(* IEC 61131-3 sources: P26002_Bosch_HDPump/P26002_Bosch_HDPump_PLC, 7 files *)

(* ---- CAN_Signals.gvl ---- *)
VAR_GLOBAL

(* ======================================================================== *)
    (* 4. Lokale Prozessvariablen für ALLE gelesenen Messwerte (Rx)             *)
    (* ======================================================================== *)
    rTecu_cpu                   : REAL; (* ID 16#456: ECU CPU Temperatur *)
    rPrail_nom                  : REAL; (* ID 16#650: Fuel pressure HP - set point *)
    rTfuel                      : REAL; (* ID 16#650: Fuel temperature HP *)
    rToil                       : REAL; (* ID 16#650: Öltemperatur *)
    rPrail_650                  : REAL; (* ID 16#650: Fuel pressure HP - side 1 *)
    rMsv_divy_angle             : REAL; (* ID 16#660: MSV Förderwinkel *)
    rAngle_eng_hdp              : REAL; (* ID 16#660: Motorwinkel HDP Messung *)
    rTinj                       : REAL; (* ID 16#660: Einspritzdauer *)
    rPrail_660                  : REAL; (* ID 16#660: Fuel pressure HP - side 2 *)
    rTekp                       : REAL; (* ID 16#670: Fuel temp after low press pump *)
    rPekp                       : REAL; (* ID 16#670: Fuel press after low press pump *)
    rPfuel                      : REAL; (* ID 16#670: Kraftstoffdruck *)
    rEngine_RPM                 : REAL; (* ID 16#680: Drehzahl / RPM *)

    (* ======================================================================== *)
    (* 5. Lokale Variablen für die zu SCHREIBENDEN Werte (Tx)                   *)
    (* ======================================================================== *)
    (* ID 16#700 *)
    rWrite_Set_RPM              : REAL  := 2500.0;
    rWrite_Actual_RPM           : REAL  := 2498.0;
    bWrite_valid_RPM            : BOOL  := TRUE;

    (* ID 16#710 *)
    rWrite_Oil_pressure         : REAL  := 4.5;    (* bar *)
    rWrite_Oil_temperature      : REAL  := 85.0;   (* °C *)
    bWrite_Oil_pressure_OK      : BOOL  := TRUE;
    bWrite_Oil_temperature_OK   : BOOL  := TRUE;

    (* ID 16#720 *)
    rWrite_Fuel_temperature     : REAL  := 25.0;   (* °C *)
    rWrite_Fuel_supply_pressure : REAL  := 5.0;    (* bar *)
    bWrite_Fuel_temperature_OK  : BOOL  := TRUE;
    bWrite_Fuel_supply_press_OK : BOOL  := TRUE;

    (* ID 16#730 *)
    rWrite_Fuel_Mass_Flow_1     : REAL  := 12.5;   (* kg/h *)
    rWrite_Fuel_Mass_Flow_2     : REAL  := 12.4;
    rWrite_Fuel_Mass_Flow_3     : REAL  := 0.0;
    bWrite_valid_Fuel_Mass_Flow : BOOL  := TRUE;

    (* ID 16#800 *)
    wWrite_ERROR_Bits           : WORD  := 16#0000;

    (* ID 16#900 *)
    nWrite_Counter_LAP          : USINT := 1;
    nWrite_Counter_FREE_TRIGGER : USINT := 0;

    (* ID 16#910 (reserviert) *)
    wWrite_RPM_Profile          : WORD  := 16#0000;

END_VAR

(* ---- GlobalVariables.gvl ---- *)
VAR_GLOBAL
system : System;
req_EmgStop_bySoftware : BOOL := FALSE;
reset_EmgStop : BOOL := FALSE;

User : User_InOut;
OP_List: ARRAY[0..10] OF OPoint;

Thermostat : Thermostat;
OilConditioning : OilConditioning;
FuelSupply : FuelSupply;

AutomaticOperation : FB_AutomaticOperation;
fbThermostat: FB_Thermostat;
fbOilConditionin: FB_OilConditioning;
fbFuelSupply: FB_FuelSupply;

HW_DI_ECU_RUNNING : BOOL; (* Kanal entsprechend benennen! *)
END_VAR

VAR_GLOBAL RETAIN
	Retain_Settings : UserSettings;
END_VAR

(* ---- FB_AutomaticOperation.st ---- *)
FUNCTION_BLOCK FB_AutomaticOperation
VAR_INPUT
	system_state : System;
	Enable  : BOOL;
    Stop    : BOOL;
    Reset   : BOOL;
    sequence_active : BOOL;

    coldStart_oil_pressure: REAL := 1.8; (* bar *)
	coldStart_oil_min_tempterature: REAL := 50; (* °C *)
	coldStart_fuelsupply_pressure: REAL := 2; (* bar *)
	coldStart_fuelsupply_min_tempterature: REAL := 50; (* °C *)
	coldStart_RPM_settings: REAL := 2000;

	normalOperation_oil_pressure: REAL := 2.5;(* bar *)
END_VAR

VAR_OUTPUT
	State   : state_op_manager; (* OP_Settle und OP_Hold brauchen wir in diesem Projekt nicht *)
    Busy    : BOOL;
    Done    : BOOL;
    Error   : BOOL;
    ErrMsg	: STRING(255);

    (* ----------------------------- *)
	(* ----- Sequence Control ------ *)
	(* ----------------------------- *)

    start_sequence: BOOL;
    stop_sequence: BOOL;
    coldStart_RPM : REAL;

     (* --- Konfiguration --- *)
    current_OP: OPoint;

END_VAR

VAR_IN_OUT
	IO_User : User_InOut;
	IO_Thermostat : Thermostat;
	IO_OilConditioning: OilConditioning;
	IO_FuelSupply: FuelSupply;
	IO_GlobalOP_List : ARRAY[0..10] OF OPoint;
END_VAR

VAR
	NextState  : state_op_manager;
    LastState  : state_op_manager;

    rpm_rampup: FB_RampTON;
    rpm_rampup_time: TIME := T#2m;
    rpm_rampup_Done: BOOL;

    prep_settle_timer: TON;
    prep_settle_time: TIME := T#60s;

	bEntry			: BOOL := TRUE;
	bInitDone       : BOOL := FALSE;
END_VAR

(* ----------------------------- *)
(* -------- Enable-Gate -------- *)
(* ----------------------------- *)
IF NOT Enable OR system_state.state = SYS_ERROR OR system_state.state = SYS_STANDBY THEN
	bInitDone := FALSE;
    State     := OP_INIT;
    LastState := OP_INIT;
    Busy      := FALSE;
    Done      := FALSE;
    Error     := FALSE;
    IO_User.Input.start := FALSE;
    RETURN;
END_IF;

(* ------------------------------------------------ *)
(* Default assignments                              *)
(* ------------------------------------------------ *)
NextState := State;
Busy  := FALSE;
Done  := FALSE;
Error := FALSE;
coldStart_RPM := 0.0;
rpm_rampup.bExecute := FALSE;
IO_Thermostat.enable := FALSE;
IO_OilConditioning.enable := FALSE;
IO_FuelSupply.enable := FALSE;

(* ------------------------------------------------ *)
(* Entry-Erkennung                                  *)
(* ------------------------------------------------ *)
bEntry := (State <> LastState);

(* ------------------------------------------------ *)
(* State Machine                                    *)
(* ------------------------------------------------ *)
CASE State OF

	OP_INIT:
	    Busy  := FALSE;
		Done  := FALSE;
		Error := FALSE;

	    IF NOT bInitDone THEN

	    ; (* Alle Infos einlesen, ggf Geräte verbinden, Geräte-Status prüfen... *)

	    bInitDone := TRUE;
	    END_IF

	    IF bInitDone THEN
	        NextState := OP_IDLE;
	        IO_User.Output.operation_status_msg := 'INFO: OP Manager initialized.';
	    END_IF

    OP_IDLE:
	    Busy  := FALSE;
		Done  := FALSE;
		Error := FALSE;

    	; (* Warten auf neue Startbedingungen *)
    	(* ------------------------------------------ *)
	    (* Startbedingung prüfen                      *)
	    (* ------------------------------------------ *)
	    Act_CheckStartConditions;

    OP_PREP:
    	Busy := TRUE;
	    Done := FALSE;
	    Error := FALSE;

	    IO_Thermostat.enable := TRUE;
		IO_OilConditioning.enable := TRUE;
		IO_FuelSupply.enable := TRUE;

	    (* Thermostat an *)
	    IO_Thermostat.target_setpoint := current_OP.Fuel_temperature;
	    IO_Thermostat.start := TRUE;

	    (* Ölkonditionierung an *)
	    IF (IO_OilConditioning.actualOil_temperature < coldStart_oil_min_tempterature+5) THEN
	    	IO_OilConditioning.setOil_pressure := coldStart_oil_pressure;
	    ELSE
	    	IF current_OP.Oil_pressure > normalOperation_oil_pressure THEN
	    		IO_OilConditioning.setOil_pressure := current_OP.Oil_pressure;
	    	ELSE
	    		IO_OilConditioning.setOil_pressure := normalOperation_oil_pressure; (* Agleich OP-Vorgabe *)
	    	END_IF
	    END_IF

	    IO_OilConditioning.setOil_temperature := current_OP.Oil_temperature; (* Wie bekomme ich die Temperatur ins ÖL? *)

	    IO_OilConditioning.start := TRUE;

	    (* Ramp up RPM *)
	    IF bEntry THEN
	    	rpm_rampup(bExecute := FALSE); (* Einmal zurücksetzen *)
	    ELSE
			rpm_rampup(
			 	bExecute := TRUE,
			 	fStartVal := 0.0,
			 	fTargetVal := coldStart_RPM_settings,
			 	tRampTime := rpm_rampup_time,
			 	fCurrentVal => coldStart_RPM,
			 	bDone => rpm_rampup_Done
			);
		END_IF

	    IF IO_Thermostat.SVreached AND
	    	IO_OilConditioning.pressure_SVreached AND
	    	IO_OilConditioning.temperature_SVreached THEN

	    	prep_settle_timer.IN := TRUE;
	    END_IF

	    IF prep_settle_timer.Q THEN
	    	IO_FuelSupply.SV := current_OP.Fuel_supply_pressure;
	    	IO_FuelSupply.start := TRUE;
	    END_IF

	    IF IO_Thermostat.SVreached AND
	    	IO_OilConditioning.pressure_SVreached AND
	    	IO_OilConditioning.temperature_SVreached AND
	    	IO_FuelSupply.SVreached AND
	    	rpm_rampup_Done THEN

	    	NextState := OP_EXECUTE;
	    END_IF

    OP_EXECUTE:
	    Busy := TRUE;
	    Done := FALSE;
	    Error := FALSE;

	    IO_Thermostat.enable := TRUE;
		IO_OilConditioning.enable := TRUE;
		IO_FuelSupply.enable := TRUE;

	    (* Benzin-Versorgung an*)
	    (* Nockenwellenantrieb nach Drehzahlvorgabe fahren*)

	OP_FINISHED:
	    Busy := FALSE;
	    Done := TRUE;
	    Error := FALSE;

	    IO_Thermostat.enable := TRUE;
		IO_OilConditioning.enable := TRUE;
(*		IO_FuelSupply.enable := TRUE; *)

	    (* Benzin-Versorgung aus *)
	    IO_FuelSupply.stop := TRUE;

	    (* Nockenwellenantrieb aus*)

	    IF IO_User.Input.continuous THEN
	    	Act_CheckStartConditions;
	    ELSE
	    	(*Cooldown: Thermostat aus, Ölkonditionierung aus*);
	    	IO_Thermostat.stop := TRUE;
	    	IO_OilConditioning.stop := TRUE;

	    END_IF

	OP_ERROR_SHUTDOWN:
	    Error := TRUE;
	    Busy := TRUE;

	OP_ERROR:
	    Error := TRUE;
	    Done := TRUE;

END_CASE;

(* ------------------------------------------------ *)
(* Global transitions                               *)
(* ------------------------------------------------ *)
IF IO_User.Input.cancel THEN
    IF State <> OP_INIT AND State <> OP_ERROR THEN
        NextState := OP_FINISHED;
        IO_User.Input.start := FALSE;
        IO_User.Input.continuous := FALSE;
    ELSIF State = OP_ERROR_SHUTDOWN THEN
    	NextState := OP_ERROR;
    	IO_User.Input.start := FALSE;
        IO_User.Input.continuous := FALSE;
    END_IF
END_IF

IF IO_User.Input.skipOP THEN
    IF State <> OP_INIT AND State <> OP_ERROR THEN
        NextState := OP_FINISHED;
        IO_User.Input.start := TRUE;
        IO_User.Input.continuous := TRUE;
    END_IF
END_IF

(* ------------------------------------------------ *)
(* ---------- Subsystem Error Detection ----------- *)
(* ------------------------------------------------ *)

(* FÜR BOSCHPRÜFSTAND: MFC FEHLER, FU Fehler, Validierungs Probleme?*)

(* IF 	(SUBP_MfcControl.ErrorDetected OR *)
(*	SUBP_HeaterControl.ErrorDetected) OR *)
(*	system.ALARM_VORALARM_H2_CT_STBQ1 AND *)
(*	State <> OP_ERROR_SHUTDOWN AND *)
(*	State <> OP_ERROR *)
(* THEN *)
(*			NextState := OP_ERROR_SHUTDOWN; *)
(*			IF SUBP_MfcControl.ErrorDetected THEN *)
(*				ErrMsg := SUBP_MfcControl.ErrMsg; *)
(*			ELSIF SUBP_HeaterControl.ErrorDetected THEN *)
(*				ErrMsg := SUBP_HeaterControl.ErrMsg; *)
(*			ELSIF system.ALARM_VORALARM_H2_CT_STBQ1 THEN *)
(*				ErrMsg := 'H2 Gas PreAlarm > 5% LowerExplosionLimit - ERROR_SHUTDOWN triggered!'; *)
(*			ELSE *)
(*				ErrMsg := 'Unknown Error detected'; *)
(*			END_IF *)
(*			Act_StateUpdate; *)
(*			RETURN; *)
(* END_IF *)

(* ------------------------------------------------ *)
(* --------- Aktualisierung Statemachine ---------- *)
(* ------------------------------------------------ *)

Act_StateUpdate;

 (* ====== PROGRAMM ENDE ====== *)
END_FUNCTION_BLOCK

ACTIONS
	ACTION Act_StateUpdate
		(* ------------------------------------------------ *)
		(* State update                                     *)
		(* ------------------------------------------------ *)
		LastState := State;
		IF NextState <> State THEN
		    State := NextState;
		END_IF;
	END_ACTION

	ACTION Act_CheckStartConditions

		current_OP := IO_GlobalOP_List[1]; (* Aktuell keine OP-Liste unterstützt *)

		IF current_OP.ProfileConfig.bDataReady AND NOT current_OP.processed THEN
			current_OP.ProfileConfig.bProfileValid := TRUE;
			NextState := OP_PREP;
		END_IF

	END_ACTION

END_ACTIONS

(* ---- MAIN.st ---- *)
PROGRAM MAIN

(*
[ ] OP_Execute
[ ] OP_Finished
[ ] FB_Thermostat
[x] FB_OilConditioning
[x] FB_FuelSupply
[ ] VERIFY RPM
[ ] VERIFY FLOW
*)
VAR
next_state : state_system;
last_state : state_system;

(* GLOBAL ERROR HANDLING *)
was_error: BOOL := FALSE;
ErrorDelayTimer : TON;         (* Delay for Error Detection *)
TriggerTime : TIME := T#1s;
ResetTrigger : TP;
StopTrigger : TP;
ALARM_ARRAY: ARRAY [1..20] OF BOOL;
a : INT; (* warnings iterative varibale *)
WARNING_ARRAY: ARRAY [1..30] OF BOOL;
w : INT; (* warnings iterative varibale *)
i : INT; (*Iteration Variable*)

(* Reset Device Errors *)
resetMfCError : BOOL;
resetEvapError : BOOL;

END_VAR

ACT_EmgStop_bySoftware;
ACT_READ_SafetyStatus;
Act_UserOutput;

ACT_StateMachine;

END_PROGRAM

ACTIONS

ACTION ACT_InitSystem
User.Settings := Retain_Settings;
;
END_ACTION

ACTION ACT_StateMachine

(* Defaults *)
AutomaticOperation.Enable := FALSE;
AutomaticOperation.Reset := FALSE;

system.state := next_state;

	CASE system.state OF
		SYS_STANDBY:
						IF system.alarm OR system.error THEN
							next_state := SYS_ERROR;
							RETURN;
						END_IF

						IF NOT system.is_init THEN
							ACT_InitSystem;
							system.is_init := TRUE;
						END_IF;

						IF User.Input.OperationModeReq THEN
							next_state := SYS_AUTO_READY;
						END_IF

		SYS_ERROR :
						ResetTrigger(IN:= User.Input.reset_Error_byUser, PT:= TriggerTime);

						IF  ResetTrigger.Q THEN
							reset_EmgStop := TRUE;
							User.Input.reset_Error_byUser := FALSE;
							AutomaticOperation.Enable := TRUE;
						END_IF

		SYS_AUTO_BUSY,SYS_AUTO_READY :

						IF system.alarm OR system.error THEN
							next_state := SYS_ERROR;
							RETURN;
						END_IF

						IF HW_DI_ECU_RUNNING THEN (* Kanal entsprechend benennen! *)
							AutomaticOperation.Enable := TRUE;
						ELSE
							AutomaticOperation.Enable := FALSE;
							 WARNING_ARRAY[2] := TRUE; (* Warnung: ECU nicht an! Kein Betrieb möglich *)
						END_IF

						IF User.Input.reset_Error_byUser THEN
							AutomaticOperation.Reset := TRUE;
						END_IF

						IF User.Input.StandbyModeReq THEN
							AutomaticOperation.Stop := TRUE;
						END_IF

		SYS_MANUAL :

						IF system.alarm OR system.error THEN
							next_state := SYS_ERROR;
							RETURN;
						END_IF

						IF User.Input.StandbyModeReq THEN
							next_state := SYS_STANDBY;
							RETURN;
						END_IF
		;
	ELSE
		next_state := SYS_ERROR; (* Other States not allowed!!! *)
		system.status_msg := 'ERROR: State Request NOT allowed!';
	END_CASE

AutomaticOperation(
 IO_User := User,
 IO_Thermostat := Thermostat,
 IO_OilConditioning := OilConditioning,
 IO_FuelSupply := FuelSupply,
 IO_GlobalOP_List := OP_List
);
fbThermostat(fbIO_Thermostat := Thermostat);
fbOilConditionin(fbIO_OilConditioning := OilConditioning);
fbFuelSupply(
 	fbIO_FuelSupply := FuelSupply,
 	SupplyFuelPumpPIDsettings := User.Settings.SupplyFuelPumpPIDsettings,
 	SupplyFuelPump_pressure_tolerance := User.Settings.SupplyFuelPump_pressure_tolerance
);

CASE AutomaticOperation.State OF

	OP_PREP, OP_EXECUTE: next_state := SYS_AUTO_BUSY;

	OP_FINISHED: next_state := SYS_STANDBY;

	OP_ERROR_SHUTDOWN, OP_ERROR: WARNING_ARRAY[1] := TRUE; (* Warnung: Automatic Programm in ERROR Condition *)

END_CASE

(* Global User Input Reset *)
User.Input.reset_Error_byUser := FALSE;
User.Input.StandbyModeReq := FALSE;
User.Input.OperationModeReq := FALSE;

last_state := system.state;
END_ACTION

ACTION Act_UserOutput

		Retain_Settings := User.Settings; (* Backup in Retain Variable *)

		User.Output.SystemState := system;

	END_ACTION

ACTION ACT_EmgStop_bySoftware
	StopTrigger(IN:= User.Input.EmgStop_Req_byUser, PT:= TriggerTime);
	req_EmgStop_bySoftware := StopTrigger.Q;

	IF req_EmgStop_bySoftware THEN
		User.Input.EmgStop_Req_byUser := FALSE;
	END_IF
	;
END_ACTION

ACTION ACT_READ_SafetyStatus (* Wird direkt im Safetyprogramm gemappt *)

		ALARM_ARRAY[1] := system.ALARM_SAI_DiagnosticError;
		ALARM_ARRAY[2] := system.ALARM_GASALARM_H2_ST_STBQ2;
		ALARM_ARRAY[3] := system.ALARM_GASALARM_H2_CT_STBQ1;
		ALARM_ARRAY[4] := system.ALARM_NotAusTaster_1_STFS1;
		ALARM_ARRAY[5] := system.ALARM_NotAusTaster_2_BPSF1;
		ALARM_ARRAY[6] := system.ALARM_EmgStop_bySoftware_activated;
		ALARM_ARRAY[7] := system.ALARM_N2Supply_STBP1;
		ALARM_ARRAY[8] := system.ALARM_HeaterLimit_T_STBT1;
		ALARM_ARRAY[9] := system.ALARM_HeaterLimit_T_STBT2;
		ALARM_ARRAY[10] := system.ALARM_NotAusTaster_1_STFS1_Discrepancy;
		ALARM_ARRAY[11] := system.ALARM_NotAusTaster_2_BPSF1_Discrepancy;
		ALARM_ARRAY[12] := system.ALARM_QA1_Discrepancy;
		ALARM_ARRAY[13] := system.ALARM_QA2_Discrepancy;
		ALARM_ARRAY[14] := system.ALARM_Draeger_Fault;

		FOR i:= 1 TO 20 DO
			IF ALARM_ARRAY[i] THEN
				system.alarm := TRUE;
			END_IF
		END_FOR

	END_ACTION

	ACTION ACT_ResetWarnings

	FOR w := 1 TO 30 DO
		WARNING_ARRAY[w] := FALSE;
	END_FOR

	END_ACTION

	ACTION ACT_CAN_COMMUNICATION
		;
	END_ACTION

END_ACTIONS

(* ---- PRG_MS7_CAN_Handler.st ---- *)
(********************************************************************************
 * PROGRAM: PRG_MS7_CAN_Handler
 *
 * Beschreibung:
 *   Erweitertes Anwendungsbeispiel für das Auslesen und Schreiben des
 *   CAN-Netzwerks (Bosch MS7 Logger / ECU) an einer Bachmann M1 Steuerung.
 *
 *   KANAL-ÜBERSICHT:
 *   ----------------------------------------------------------------------------
 *   EMPFANG (R / Rx):
 *     - Kanal 1 (Rx): ID 16#650 (prail_nom, tfuel, toil, prail_650)
 *     - Kanal 2 (Rx): ID 16#660 (msv_divy_angle, angle_eng_hdp, tinj, prail_660)
 *     - Kanal 3 (Rx): ID 16#670 (tEKP, pEKP, pfuel)
 *     - Kanal 4 (Rx): ID 16#456 (tecu_cpu)
 *     - Kanal 5 (Rx): ID 16#680 (Drehzahl / RPM)
 *
 *   SENDEN (W / Tx):
 *     - Kanal 6  (Tx): ID 16#700 (Set RPM, Actual RPM, valid RPM)
 *     - Kanal 7  (Tx): ID 16#710 (Oil pressure, Oil temperature, Status OK-Bits)
 *     - Kanal 8  (Tx): ID 16#720 (Fuel temp, Fuel supply press, Status OK-Bits)
 *     - Kanal 9  (Tx): ID 16#730 (Fuel Mass Flow 1, 2, 3, valid Bit)
 *     - Kanal 10 (Tx): ID 16#800 (ERROR_Bits)
 *     - Kanal 11 (Tx): ID 16#900 (Counter LAP, Counter FREE TRIGGER)
 *     - Kanal 12 (Tx): ID 16#910 (RPM Profile - reserviert)
 ********************************************************************************)
PROGRAM PRG_MS7_CAN_Handler
VAR
    (* ======================================================================== *)
    (* 1. Konfigurationstabelle / Maske aller CAN-Kanäle (Botschaftsebene)      *)
    (* ======================================================================== *)
    canChannels                 : ARRAY [1..32] OF ST_CAN_Broker_Channel;
    bConfigDone                 : BOOL := FALSE;

    (* Hardware CAN-Broker Instanz (modular bis 32 Kanäle) *)
    fbBroker                    : FB_CAN_Broker_Modular;
    bBrokerReady                : BOOL;
    bBrokerError                : BOOL;
    nBrokerErrorID              : DINT;

    (* ======================================================================== *)
    (* 2. Signal-Instanzen zum LESEN (Rx)                                       *)
    (* ======================================================================== *)
    (* Kanal 4: Botschaft 16#456 (1110 dez) *)
    fb_tecu_cpu                 : FB_CAN_Signal;

    (* Kanal 1: Botschaft 16#650 (1616 dez) *)
    fb_prail_nom                : FB_CAN_Signal; (* Fuel press HP - set point (Bit 0, 16 Bit) *)
    fb_tfuel                    : FB_CAN_Signal; (* Fuel temp HP (Bit 16, 8 Bit) *)
    fb_toil                     : FB_CAN_Signal; (* Oil temp (Bit 24, 8 Bit) *)
    fb_prail_650                : FB_CAN_Signal; (* Fuel press HP - side 1 (Bit 48, 16 Bit) *)

    (* Kanal 2: Botschaft 16#660 (1632 dez) *)
    fb_msv_divy_angle           : FB_CAN_Signal;
    fb_angle_eng_hdp            : FB_CAN_Signal;
    fb_tinj                     : FB_CAN_Signal;
    fb_prail_660                : FB_CAN_Signal; (* Fuel press HP - side 2 (Bit 48, 16 Bit) *)

    (* Kanal 3: Botschaft 16#670 (1648 dez) *)
    fb_tEKP                     : FB_CAN_Signal; (* Fuel temp after low press pump (Bit 0, 16 Bit) *)
    fb_pEKP                     : FB_CAN_Signal; (* Fuel press after low press pump (Bit 16, 16 Bit) *)
    fb_pfuel                    : FB_CAN_Signal; (* Fuel pressure (Bit 32, 8 Bit) *)

    (* Kanal 5: Botschaft 16#680 (1664 dez) *)
    fb_engine_RPM               : FB_CAN_Signal; (* Drehzahl / RPM (Bit 0, 16 Bit) *)

    (* ======================================================================== *)
    (* 3. Signal-Instanzen zum SCHREIBEN (Tx)                                   *)
    (* ======================================================================== *)
    (* Kanal 6: Botschaft 16#700 (1792 dez) *)
    fb_w_Set_RPM                : FB_CAN_Signal; (* Set RPM (Bit 0, 16 Bit) *)
    fb_w_Actual_RPM             : FB_CAN_Signal; (* Actual RPM (Bit 16, 16 Bit) *)
    fb_w_valid_RPM              : FB_CAN_Signal; (* valid RPM (Bit 32, 16 Bit) *)

    (* Kanal 7: Botschaft 16#710 (1808 dez) *)
    fb_w_Oil_pressure           : FB_CAN_Signal; (* Oil pressure (Bit 0, 16 Bit) *)
    fb_w_Oil_temperature        : FB_CAN_Signal; (* Oil temperature (Bit 16, 16 Bit) *)
    fb_w_Oil_pressure_OK        : FB_CAN_Signal; (* Oil pressure OK (Bit 32, 1 Bit) *)
    fb_w_Oil_temperature_OK     : FB_CAN_Signal; (* Oil temperature OK (Bit 33, 1 Bit) *)

    (* Kanal 8: Botschaft 16#720 (1824 dez) *)
    fb_w_Fuel_temperature       : FB_CAN_Signal; (* Fuel temperature (Bit 0, 16 Bit) *)
    fb_w_Fuel_supply_pressure   : FB_CAN_Signal; (* Fuel supply pressure (Bit 16, 16 Bit) *)
    fb_w_Fuel_temperature_OK    : FB_CAN_Signal; (* Fuel temperature OK (Bit 32, 1 Bit) *)
    fb_w_Fuel_supply_press_OK   : FB_CAN_Signal; (* Fuel supply pressure OK (Bit 33, 1 Bit) *)

    (* Kanal 9: Botschaft 16#730 (1840 dez) *)
    fb_w_Fuel_Mass_Flow_1       : FB_CAN_Signal; (* Fuel Mass Flow 1 (Bit 0, 16 Bit) *)
    fb_w_Fuel_Mass_Flow_2       : FB_CAN_Signal; (* Fuel Mass Flow 2 (Bit 16, 16 Bit) *)
    fb_w_Fuel_Mass_Flow_3       : FB_CAN_Signal; (* Fuel Mass Flow 3 (Bit 32, 16 Bit) *)
    fb_w_valid_Fuel_Mass_Flow   : FB_CAN_Signal; (* valid Fuel Mass Flow (Bit 48, 1 Bit) *)

    (* Kanal 10: Botschaft 16#800 (2048 dez) *)
    fb_w_ERROR_Bits             : FB_CAN_Signal; (* ERROR_Bits (Bit 0, 16 Bit) *)

    (* Kanal 11: Botschaft 16#900 (2304 dez) *)
    fb_w_Counter_LAP            : FB_CAN_Signal; (* Counter Byte 1 (LAP) (Bit 0, 8 Bit) *)
    fb_w_Counter_FREE_TRIGGER   : FB_CAN_Signal; (* Counter Byte 2 (FREE TRIGGER) (Bit 8, 8 Bit) *)

    (* Kanal 12: Botschaft 16#910 (2320 dez) *)
    fb_w_RPM_Profile            : FB_CAN_Signal; (* RPM Profile (reserviert) *)

(*     (* ======================================================================== *) *)
(*     (* 4. Lokale Prozessvariablen für ALLE gelesenen Messwerte (Rx)             *) *)
(*     (* ======================================================================== *) *)
(*     rTecu_cpu                   : REAL; (* ID 16#456: ECU CPU Temperatur *) *)
(*     rPrail_nom                  : REAL; (* ID 16#650: Fuel pressure HP - set point *) *)
(*     rTfuel                      : REAL; (* ID 16#650: Fuel temperature HP *) *)
(*     rToil                       : REAL; (* ID 16#650: Öltemperatur *) *)
(*     rPrail_650                  : REAL; (* ID 16#650: Fuel pressure HP - side 1 *) *)
(*     rMsv_divy_angle             : REAL; (* ID 16#660: MSV Förderwinkel *) *)
(*     rAngle_eng_hdp              : REAL; (* ID 16#660: Motorwinkel HDP Messung *) *)
(*     rTinj                       : REAL; (* ID 16#660: Einspritzdauer *) *)
(*     rPrail_660                  : REAL; (* ID 16#660: Fuel pressure HP - side 2 *) *)
(*     rTekp                       : REAL; (* ID 16#670: Fuel temp after low press pump *) *)
(*     rPekp                       : REAL; (* ID 16#670: Fuel press after low press pump *) *)
(*     rPfuel                      : REAL; (* ID 16#670: Kraftstoffdruck *) *)
(*     rEngine_RPM                 : REAL; (* ID 16#680: Drehzahl / RPM *) *)
(*  *)
(*     (* ======================================================================== *) *)
(*     (* 5. Lokale Variablen für die zu SCHREIBENDEN Werte (Tx)                   *) *)
(*     (* ======================================================================== *) *)
(*     (* ID 16#700 *) *)
(*     rWrite_Set_RPM              : REAL  := 2500.0; *)
(*     rWrite_Actual_RPM           : REAL  := 2498.0; *)
(*     bWrite_valid_RPM            : BOOL  := TRUE; *)
(*  *)
(*     (* ID 16#710 *) *)
(*     rWrite_Oil_pressure         : REAL  := 4.5;    (* bar *) *)
(*     rWrite_Oil_temperature      : REAL  := 85.0;   (* °C *) *)
(*     bWrite_Oil_pressure_OK      : BOOL  := TRUE; *)
(*     bWrite_Oil_temperature_OK   : BOOL  := TRUE; *)
(*  *)
(*     (* ID 16#720 *) *)
(*     rWrite_Fuel_temperature     : REAL  := 25.0;   (* °C *) *)
(*     rWrite_Fuel_supply_pressure : REAL  := 5.0;    (* bar *) *)
(*     bWrite_Fuel_temperature_OK  : BOOL  := TRUE; *)
(*     bWrite_Fuel_supply_press_OK : BOOL  := TRUE; *)
(*  *)
(*     (* ID 16#730 *) *)
(*     rWrite_Fuel_Mass_Flow_1     : REAL  := 12.5;   (* kg/h *) *)
(*     rWrite_Fuel_Mass_Flow_2     : REAL  := 12.4; *)
(*     rWrite_Fuel_Mass_Flow_3     : REAL  := 0.0; *)
(*     bWrite_valid_Fuel_Mass_Flow : BOOL  := TRUE; *)
(*  *)
(*     (* ID 16#800 *) *)
(*     wWrite_ERROR_Bits           : WORD  := 16#0000; *)
(*  *)
(*     (* ID 16#900 *) *)
(*     nWrite_Counter_LAP          : USINT := 1; *)
(*     nWrite_Counter_FREE_TRIGGER : USINT := 0; *)
(*  *)
(*     (* ID 16#910 (reserviert) *) *)
(*     wWrite_RPM_Profile          : WORD  := 16#0000; *)

    (* ======================================================================== *)
    (* 6. Sende-Steuerung (Zykluszähler für 10 ms Task -> 100 ms Takt)         *)
    (* ======================================================================== *)
    bContinuousSend             : BOOL := TRUE;      (* TRUE = Kontinuierlich alle 100 ms senden *)
    nCycleCounter               : INT  := 0;         (* Zykluszähler *)
    nTargetCycles               : INT  := 10;        (* 10 Zyklen à 10 ms = exakt 100.0 ms *)
    bSendTriggerManual          : BOOL := FALSE;     (* Manueller Einzeltakt-Trigger *)

    (* Einzelne Sende-Freigaben für jede Botschaft *)
    bEnableTx_700               : BOOL := TRUE;
    bEnableTx_710               : BOOL := TRUE;
    bEnableTx_720               : BOOL := TRUE;
    bEnableTx_730               : BOOL := TRUE;
    bEnableTx_800               : BOOL := TRUE;
    bEnableTx_900               : BOOL := TRUE;
    bEnableTx_910               : BOOL := FALSE;     (* Reserviert - Standard inaktiv *)
END_VAR

(* ============================================================================ *)
(* Initialisierung der Kanal-Maske (1..12)                                      *)
(* ============================================================================ *)
IF NOT bConfigDone THEN
    (* Empfangskanäle (Rx) *)
    canChannels[1].RxCobId := 16#650;  canChannels[1].TxCobId := 0;
    canChannels[2].RxCobId := 16#660;  canChannels[2].TxCobId := 0;
    canChannels[3].RxCobId := 16#670;  canChannels[3].TxCobId := 0;
    canChannels[4].RxCobId := 16#456;  canChannels[4].TxCobId := 0;
    canChannels[5].RxCobId := 16#680;  canChannels[5].TxCobId := 0;

    (* Sendekanäle (Tx) *)
    canChannels[6].TxCobId  := 16#700; canChannels[6].RxCobId  := 0;
    canChannels[7].TxCobId  := 16#710; canChannels[7].RxCobId  := 0;
    canChannels[8].TxCobId  := 16#720; canChannels[8].RxCobId  := 0;
    canChannels[9].TxCobId  := 16#730; canChannels[9].RxCobId  := 0;
    canChannels[10].TxCobId := 16#800; canChannels[10].RxCobId := 0;
    canChannels[11].TxCobId := 16#900; canChannels[11].RxCobId := 0;
    canChannels[12].TxCobId := 16#910; canChannels[12].RxCobId := 0;

    bConfigDone := TRUE;
END_IF;

(* ============================================================================ *)
(* 1. Hardware CAN-Broker aufrufen (NumChannels := 12)                          *)
(* ============================================================================ *)
fbBroker(
    Enable      := TRUE,
    Reset       := FALSE,
    NetNb       := 1,
    CardNb      := 2,
    Chan        := 0,
    NumChannels := 12,
    Channels    := canChannels,
    Ready       => bBrokerReady,
    Error       => bBrokerError,
    ErrorID     => nBrokerErrorID
);

(* ============================================================================ *)
(* 2. EMPFANGEN (Rx): Signale decodieren                                        *)
(* ============================================================================ *)

(* Kanal 4: ID 16#456 (tecu_cpu) *)
fb_tecu_cpu(
    CobId     := 16#456,
    StartBit  := 0,
    BitLength := 16,
    bWrite    := FALSE,
    Data      := canChannels[4].RxData
);
rTecu_cpu := fb_tecu_cpu.PhysValue;

(* Kanal 1: ID 16#650 *)
fb_prail_nom(
    CobId     := 16#650,
    StartBit  := 0,
    BitLength := 16,
    bWrite    := FALSE,
    Data      := canChannels[1].RxData
);
rPrail_nom := fb_prail_nom.PhysValue;

fb_tfuel(
    CobId     := 16#650,
    StartBit  := 16,
    BitLength := 8,
    bWrite    := FALSE,
    Data      := canChannels[1].RxData
);
rTfuel := fb_tfuel.PhysValue;

fb_toil(
    CobId     := 16#650,
    StartBit  := 24,
    BitLength := 8,
    bWrite    := FALSE,
    Data      := canChannels[1].RxData
);
rToil := fb_toil.PhysValue;

fb_prail_650(
    CobId     := 16#650,
    StartBit  := 48,
    BitLength := 16,
    bWrite    := FALSE,
    Data      := canChannels[1].RxData
);
rPrail_650 := fb_prail_650.PhysValue;

(* Kanal 2: ID 16#660 *)
fb_msv_divy_angle(
    CobId     := 16#660,
    StartBit  := 0,
    BitLength := 16,
    bWrite    := FALSE,
    Data      := canChannels[2].RxData
);
rMsv_divy_angle := fb_msv_divy_angle.PhysValue;

fb_angle_eng_hdp(
    CobId     := 16#660,
    StartBit  := 16,
    BitLength := 16,
    bWrite    := FALSE,
    Data      := canChannels[2].RxData
);
rAngle_eng_hdp := fb_angle_eng_hdp.PhysValue;

fb_tinj(
    CobId     := 16#660,
    StartBit  := 32,
    BitLength := 16,
    bWrite    := FALSE,
    Data      := canChannels[2].RxData
);
rTinj := fb_tinj.PhysValue;

fb_prail_660(
    CobId     := 16#660,
    StartBit  := 48,
    BitLength := 16,
    bWrite    := FALSE,
    Data      := canChannels[2].RxData
);
rPrail_660 := fb_prail_660.PhysValue;

(* Kanal 3: ID 16#670 *)
fb_tEKP(
    CobId     := 16#670,
    StartBit  := 0,
    BitLength := 16,
    bWrite    := FALSE,
    Data      := canChannels[3].RxData
);
rTekp := fb_tEKP.PhysValue;

fb_pEKP(
    CobId     := 16#670,
    StartBit  := 16,
    BitLength := 16,
    bWrite    := FALSE,
    Data      := canChannels[3].RxData
);
rPekp := fb_pEKP.PhysValue;

fb_pfuel(
    CobId     := 16#670,
    StartBit  := 32,
    BitLength := 8,
    bWrite    := FALSE,
    Data      := canChannels[3].RxData
);
rPfuel := fb_pfuel.PhysValue;

(* Kanal 5: ID 16#680 (Drehzahl / RPM) *)
fb_engine_RPM(
    CobId     := 16#680,
    StartBit  := 0,
    BitLength := 16,
    bWrite    := FALSE,
    Data      := canChannels[5].RxData
);
rEngine_RPM := fb_engine_RPM.PhysValue;

(* ============================================================================ *)
(* 3. SENDEN (Tx): Botschaften packen und alle 100 ms an Broker übergeben       *)
(* ============================================================================ *)
IF bContinuousSend THEN
    nCycleCounter := nCycleCounter + 1;
END_IF;

(* Senden auslösen: Exakt bei jedem 10. SPS-Durchlauf (100 ms) oder per Trigger *)
IF ((bContinuousSend AND (nCycleCounter >= nTargetCycles)) OR bSendTriggerManual) THEN

    nCycleCounter := 0; (* Zähler zurücksetzen *)

    (* ------------------------------------------------------------------------ *)
    (* Kanal 6: ID 16#700 (Set RPM, Actual RPM, valid RPM)                      *)
    (* ------------------------------------------------------------------------ *)
    IF bEnableTx_700 AND NOT canChannels[6].TxBusy THEN
        fb_w_Set_RPM(
            CobId      := 16#700,
            StartBit   := 0,
            BitLength  := 16,
            bWrite     := TRUE,
            WriteValue := rWrite_Set_RPM,
            Data       := canChannels[6].TxData
        );
        fb_w_Actual_RPM(
            CobId      := 16#700,
            StartBit   := 16,
            BitLength  := 16,
            bWrite     := TRUE,
            WriteValue := rWrite_Actual_RPM,
            Data       := canChannels[6].TxData
        );
        fb_w_valid_RPM(
            CobId      := 16#700,
            StartBit   := 32,
            BitLength  := 16,
            bWrite     := TRUE,
            WriteValue := SEL(bWrite_valid_RPM, 0.0, 1.0),
            Data       := canChannels[6].TxData
        );
        canChannels[6].TxReq := TRUE;
    END_IF;

    (* ------------------------------------------------------------------------ *)
    (* Kanal 7: ID 16#710 (Oil pressure, Oil temperature, Status OK-Bits)       *)
    (* ------------------------------------------------------------------------ *)
    IF bEnableTx_710 AND NOT canChannels[7].TxBusy THEN
        fb_w_Oil_pressure(
            CobId      := 16#710,
            StartBit   := 0,
            BitLength  := 16,
            bWrite     := TRUE,
            WriteValue := rWrite_Oil_pressure,
            Data       := canChannels[7].TxData
        );
        fb_w_Oil_temperature(
            CobId      := 16#710,
            StartBit   := 16,
            BitLength  := 16,
            bWrite     := TRUE,
            WriteValue := rWrite_Oil_temperature,
            Data       := canChannels[7].TxData
        );
        fb_w_Oil_pressure_OK(
            CobId      := 16#710,
            StartBit   := 32,
            BitLength  := 1,
            bWrite     := TRUE,
            WriteValue := SEL(bWrite_Oil_pressure_OK, 0.0, 1.0),
            Data       := canChannels[7].TxData
        );
        fb_w_Oil_temperature_OK(
            CobId      := 16#710,
            StartBit   := 33,
            BitLength  := 1,
            bWrite     := TRUE,
            WriteValue := SEL(bWrite_Oil_temperature_OK, 0.0, 1.0),
            Data       := canChannels[7].TxData
        );
        canChannels[7].TxReq := TRUE;
    END_IF;

    (* ------------------------------------------------------------------------ *)
    (* Kanal 8: ID 16#720 (Fuel temp, Fuel supply press, Status OK-Bits)        *)
    (* ------------------------------------------------------------------------ *)
    IF bEnableTx_720 AND NOT canChannels[8].TxBusy THEN
        fb_w_Fuel_temperature(
            CobId      := 16#720,
            StartBit   := 0,
            BitLength  := 16,
            bWrite     := TRUE,
            WriteValue := rWrite_Fuel_temperature,
            Data       := canChannels[8].TxData
        );
        fb_w_Fuel_supply_pressure(
            CobId      := 16#720,
            StartBit   := 16,
            BitLength  := 16,
            bWrite     := TRUE,
            WriteValue := rWrite_Fuel_supply_pressure,
            Data       := canChannels[8].TxData
        );
        fb_w_Fuel_temperature_OK(
            CobId      := 16#720,
            StartBit   := 32,
            BitLength  := 1,
            bWrite     := TRUE,
            WriteValue := SEL(bWrite_Fuel_temperature_OK, 0.0, 1.0),
            Data       := canChannels[8].TxData
        );
        fb_w_Fuel_supply_press_OK(
            CobId      := 16#720,
            StartBit   := 33,
            BitLength  := 1,
            bWrite     := TRUE,
            WriteValue := SEL(bWrite_Fuel_supply_press_OK, 0.0, 1.0),
            Data       := canChannels[8].TxData
        );
        canChannels[8].TxReq := TRUE;
    END_IF;

    (* ------------------------------------------------------------------------ *)
    (* Kanal 9: ID 16#730 (Fuel Mass Flow 1, 2, 3, valid Bit)                   *)
    (* ------------------------------------------------------------------------ *)
    IF bEnableTx_730 AND NOT canChannels[9].TxBusy THEN
        fb_w_Fuel_Mass_Flow_1(
            CobId      := 16#730,
            StartBit   := 0,
            BitLength  := 16,
            bWrite     := TRUE,
            WriteValue := rWrite_Fuel_Mass_Flow_1,
            Data       := canChannels[9].TxData
        );
        fb_w_Fuel_Mass_Flow_2(
            CobId      := 16#730,
            StartBit   := 16,
            BitLength  := 16,
            bWrite     := TRUE,
            WriteValue := rWrite_Fuel_Mass_Flow_2,
            Data       := canChannels[9].TxData
        );
        fb_w_Fuel_Mass_Flow_3(
            CobId      := 16#730,
            StartBit   := 32,
            BitLength  := 16,
            bWrite     := TRUE,
            WriteValue := rWrite_Fuel_Mass_Flow_3,
            Data       := canChannels[9].TxData
        );
        fb_w_valid_Fuel_Mass_Flow(
            CobId      := 16#730,
            StartBit   := 48,
            BitLength  := 1,
            bWrite     := TRUE,
            WriteValue := SEL(bWrite_valid_Fuel_Mass_Flow, 0.0, 1.0),
            Data       := canChannels[9].TxData
        );
        canChannels[9].TxReq := TRUE;
    END_IF;

    (* ------------------------------------------------------------------------ *)
    (* Kanal 10: ID 16#800 (ERROR_Bits)                                         *)
    (* ------------------------------------------------------------------------ *)
    IF bEnableTx_800 AND NOT canChannels[10].TxBusy THEN
        fb_w_ERROR_Bits(
            CobId      := 16#800,
            StartBit   := 0,
            BitLength  := 16,
            bWrite     := TRUE,
            WriteValue := DINT_TO_REAL(WORD_TO_DINT(wWrite_ERROR_Bits)),
            Data       := canChannels[10].TxData
        );
        canChannels[10].TxReq := TRUE;
    END_IF;

    (* ------------------------------------------------------------------------ *)
    (* Kanal 11: ID 16#900 (Counter LAP, Counter FREE TRIGGER)                  *)
    (* ------------------------------------------------------------------------ *)
    IF bEnableTx_900 AND NOT canChannels[11].TxBusy THEN
        fb_w_Counter_LAP(
            CobId      := 16#900,
            StartBit   := 0,
            BitLength  := 8,
            bWrite     := TRUE,
            WriteValue := USINT_TO_REAL(nWrite_Counter_LAP),
            Data       := canChannels[11].TxData
        );
        fb_w_Counter_FREE_TRIGGER(
            CobId      := 16#900,
            StartBit   := 8,
            BitLength  := 8,
            bWrite     := TRUE,
            WriteValue := USINT_TO_REAL(nWrite_Counter_FREE_TRIGGER),
            Data       := canChannels[11].TxData
        );
        canChannels[11].TxReq := TRUE;
    END_IF;

    (* ------------------------------------------------------------------------ *)
    (* Kanal 12: ID 16#910 (RPM Profile - reserviert)                           *)
    (* ------------------------------------------------------------------------ *)
    IF bEnableTx_910 AND NOT canChannels[12].TxBusy THEN
        fb_w_RPM_Profile(
            CobId      := 16#910,
            StartBit   := 0,
            BitLength  := 16,
            bWrite     := TRUE,
            WriteValue := DINT_TO_REAL(WORD_TO_DINT(wWrite_RPM_Profile)),
            Data       := canChannels[12].TxData
        );
        canChannels[12].TxReq := TRUE;
    END_IF;

    bSendTriggerManual := FALSE;

END_IF;

END_PROGRAM

(* ---- PRG_RPM_Control_1ms.st ---- *)
(********************************************************************************
 * PROGRAM: PRG_RPM_Control_1ms
 *
 * Beschreibung:
 *   Hauptprogramm für die Motoransteuerung im 1-ms-Echtzeittask.
 *   - Umschaltbar zwischen:
 *       0 = Dreiecksprofil (FB_TriangleProfile)
 *       1 = Sinusprofil mit Phasenversatz (FB_SineProfile)
 *       2 = 10-ms-OPC-UA-Profil (FB_ArrayProfile)
 *   - Sequenzüberwachung mit Zähler- und 48h-Zeitabschaltung
 *   - bSequenceActiveOut (Start/End-Signal) & bLapTriggerOut (gepulst)
 *   - Profibus-Telegrammausgabe an den Frequenzumrichter
 ********************************************************************************)
PROGRAM PRG_RPM_Control_1ms
VAR

    (* --- Konfiguration --- *)
    fRampAccelPreset    : REAL              := 500.0; (* U/s Beschleunigung *)

    (* --- Bedienung & Status --- *)
    bLapTriggerOut      : BOOL;
    fTargetRpm			: REAL;
    bCmdResetDrive      : BOOL;
    bDriveReadyOut      : BOOL;
    bDriveErrorOut      : BOOL;

    (* --- Baustein-Instanzen --- *)
    fbSeq               : FB_SequenceController;
    fbTriangle          : FB_TriangleProfile;
    fbSine              : FB_SineProfile;
    fbArrayPlayer       : FB_ArrayProfile;
    fbDrive             : FB_ProfibusDrive;

    (* --- Interne Signale --- *)
    fCurrentRpm         : REAL;
    fActualRpmNW        : REAL;
    bLapSignal          : BOOL;

    (* --- PROFINET / PROFIBUS I/O Mapping (Slot 4: SEW MOVIAXIS) --- *)
    (* Ausgänge an Umrichter (PA 1..4 = 8 Byte) *)
(*     q_SEW_Action        AT %Q* : INT;   (* PA 1: Aktion (20 = Linkslauf, 32 = Reset, 0 = Stopp) *) *)
(*     q_SEW_SpeedSetpoint AT %Q* : INT;   (* PA 2: Motordrehzahl = Nockenwellendrehzahl / 1.43 *) *)
(*     q_SEW_Accel         AT %Q* : INT;   (* PA 3: Beschleunigung [U/s] *) *)
(*     q_SEW_Ruck          AT %Q* : INT;   (* PA 4: Ruck (fest 0) *) *)
(*  *)
(*     (* Eingänge von Umrichter (PE 1..4 = 8 Byte) *) *)
(*     i_SEW_StatusWord    AT %I* : WORD;  (* PE 1: Statuswort Umrichter *) *)
(*     i_SEW_ActualSpeed   AT %I* : INT;   (* PE 2: Motor-Istdrehzahl *) *)
(*     i_SEW_ActualCurrent AT %I* : INT;   (* PE 3: Motorstrom *) *)
(*     i_SEW_DiagInfo      AT %I* : WORD;  (* PE 4: Diagnose / Fehlercode *) *)
END_VAR

(* 1. Profilberechnung je nach Auswahl *)
CASE AutomaticOperation.current_OP.ProfileType OF
    PROFILE_TRIANGLE:
        fbTriangle(
            bExecute     := fbSeq.bSequenceActive,
            stConfig     := AutomaticOperation.current_OP.ProfileConfig.TriangleConfig,
            tCycleTime   := T#1ms,
            fRpmOut      => fCurrentRpm,
            bLapFinished => bLapSignal
        );

    PROFILE_SINE:
        fbSine(
            bExecute     := fbSeq.bSequenceActive,
            stConfig     := AutomaticOperation.current_OP.ProfileConfig.SineConfig,
            tCycleTime   := T#1ms,
            fRpmOut      => fCurrentRpm,
            bLapFinished => bLapSignal
        );

    PROFILE_ARRAY_10MS:
        fbArrayPlayer(
            bExecute       := fbSeq.bSequenceActive,
            nPointsInLap   := AutomaticOperation.current_OP.ProfileConfig.FreeConfig.nPointsCount,
            aLapDataBuffer := AutomaticOperation.current_OP.ProfileConfig.FreeConfig.LapData,
            fRpmOut        => fCurrentRpm,
            bLapFinished   => bLapSignal
        );
END_CASE;

(* 2. Sequenz-Controller *)
fbSeq(
    bStart              := AutomaticOperation.start_sequence,
    bStop               := AutomaticOperation.stop_sequence,
    eEndMode            := AutomaticOperation.current_OP.ProfileConfig.eEndMode,
    nTargetLaps         := AutomaticOperation.current_OP.ProfileConfig.nLaps,
    tTargetDuration     := AutomaticOperation.current_OP.ProfileConfig.tDuration,
    tLapPulseDuration   := User.Settings.tLapPulseLen,
    bLapFinishedSignal  := bLapSignal,
    tCycleTime          := T#1ms,
    bSequenceActive     => AutomaticOperation.sequence_active,
    bLapTrigger         => bLapTriggerOut,
    nCompletedLaps      => User.Output.nActualLaps,       (* <- HIER: Rundenanzahl abholen *)
    tElapsedTime        => User.Output.tActualTime        (* <- HIER: Bisherige Laufzeit abholen *)
);

(* 3. Ausgabe an Frequenzumrichter *)
IF AutomaticOperation.State = OP_PREP THEN
	fTargetRpm := AutomaticOperation.coldStart_RPM;
	fbDrive.bEnable := TRUE;
ELSIF fbSeq.bSequenceActive THEN
	fTargetRpm := fCurrentRpm;
	fbDrive.bEnable := TRUE;
ELSE (* Wenn Sequenz AUS ist: Solldrehzahl GARANTIERT auf 0.0 zwingen! *)
	fTargetRpm := 0.0;
	fbDrive.bEnable := FALSE;
END_IF

fbDrive(
    bReset              := bCmdResetDrive,
    bDirectionReverse   := FALSE, (* FALSE = Linkslauf (HDP-Standard) *)
    fRpmSetpoint   		:= fTargetRpm,
    fRampAccel          := fRampAccelPreset,
    fGearRatio          := 1.43,
(*     i_nStatusWord       := i_SEW_StatusWord, *)
(*     i_nActualSpeed      := i_SEW_ActualSpeed, *)
(*     i_nActualCurrent    := i_SEW_ActualCurrent, *)
(*     i_nDiagInfo         := i_SEW_DiagInfo, *)
(*     q_nActionCode       => q_SEW_Action, *)
(*     q_nSpeedSetpoint    => q_SEW_SpeedSetpoint, *)
(*     q_nRampAccel        => q_SEW_Accel, *)
(*     q_nRuck             => q_SEW_Ruck, *)
    rActualRpmNW        => fActualRpmNW,
    bDriveReady         => bDriveReadyOut,
    bDriveError         => bDriveErrorOut
);

END_PROGRAM

(* ---- SUBP_SignalLights.st ---- *)
PROGRAM SUBP_SignalLights
VAR

END_VAR

ACT_StateLights;
(* SUBP_HWmapping_Lights; *) (* KEINE HW vorhanden*)

END_PROGRAM

ACTIONS
(* Bedienpanel: alles gleiche Schriftgröße *)
(*	- NOT-Aus --> NOT-Aus *)
(*	- rot --> Alarm \ Reset *)
(*	- gelb --> Betrieb \ Start *)
(*	- grün --> Stand-BY \ Stop *)
(*	ggf. vor Befehl Symbole setzen (Lampe + Hand o.Ä.) *)
(*	Kommentare Lukas: *)
(*		Symbole vor den Text wären sinnvoll *)
(*		rot --> Alarm / Reset (damit sind Anzeige und Funktionalität auf einem Leuchttaster) *)
(*			konstant: Warnung *)
(*			blinkend: Alarm *)
(*		gelb --> Betrieb / Start - startet eine vordefinierte Sequenz im Automatikmodus *)
(*			konstant: Betrieb - Eingeregelt *)
(*			blinkend: Betrieb - transient oder Manueller Modus *)
(*		grün --> Standby / Softstop - In den Standby fahren, inkl CoolDown und N2-Spülen  *)
(*			konstant: Alles sicher, Prüfstand tut nix *)
(*			blinkend: Heizungen / Ventile bestromt *)

	 ACTION ACT_StateLights
	 	CASE system.state OF

	    1: (* ERROR *)

	        User.Output.Ampel_rot := TRUE;
	        User.Output.Ampel_rot_blink := FALSE;
	        User.Output.Ampel_gelb := FALSE;
	        User.Output.Ampel_gelb_blink := FALSE;
	        User.Output.Ampel_gruen := FALSE;
	        User.Output.Ampel_gruen_blink := FALSE;

	    0: (* Standby *)

	    	User.Output.Ampel_rot := FALSE;
	        User.Output.Ampel_rot_blink := FALSE;
	        User.Output.Ampel_gelb := FALSE;
	        User.Output.Ampel_gelb_blink := FALSE;
	        User.Output.Ampel_gruen := TRUE;
	        User.Output.Ampel_gruen_blink := FALSE;

	    2,3: (* Automatic *)
	    	CASE AutomaticOperation.State OF
	    		OP_INIT,OP_IDLE:

							        User.Output.Ampel_rot := FALSE;
							        User.Output.Ampel_rot_blink := FALSE;
							        User.Output.Ampel_gelb := FALSE;
							        User.Output.Ampel_gelb_blink := FALSE;
							        User.Output.Ampel_gruen := FALSE;
							        User.Output.Ampel_gruen_blink := TRUE;

		    	OP_HOLD,OP_FINISHED:

							        User.Output.Ampel_rot := FALSE;
							        User.Output.Ampel_rot_blink := FALSE;
							        User.Output.Ampel_gelb := TRUE;
							        User.Output.Ampel_gelb_blink := FALSE;
							        User.Output.Ampel_gruen := FALSE;
							        User.Output.Ampel_gruen_blink := FALSE;

			    OP_PREP, OP_EXECUTE, OP_WAIT_SETTLED:

							        User.Output.Ampel_rot := FALSE;
							        User.Output.Ampel_rot_blink := FALSE;
							        User.Output.Ampel_gelb := FALSE;
							        User.Output.Ampel_gelb_blink := TRUE;
							        User.Output.Ampel_gruen := FALSE;
							        User.Output.Ampel_gruen_blink := FALSE;
		    END_CASE

	    4: (* Manual Operation Mode *)

	        User.Output.Ampel_rot := FALSE;
	        User.Output.Ampel_rot_blink := FALSE;
	        User.Output.Ampel_gelb := FALSE;
	        User.Output.Ampel_gelb_blink := TRUE;
	        User.Output.Ampel_gruen := FALSE;
	        User.Output.Ampel_gruen_blink := FALSE;

		END_CASE

		IF system.state <> 1 AND system.warning THEN
			User.Output.Ampel_rot_blink := TRUE;
		END_IF
	 END_ACTION

END_ACTIONS
